FUNCTION_BLOCK MOD_StateLatch (* Keeps the last module state heard on the state channel. Technical: Local channel IDs of the PackML state and its refresh query; types and forwards the received PackML state *)
  (* Standard: 61499-2 *)
  (* Version 0.1, 2026-09-28, Project contributors, AAU Smart Production Lab *)
  PACKAGE modlib;
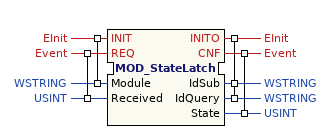
  EVENT_INPUT
    INIT : EInit WITH Module; (* Initialise, once at start-up (the INIT chain); takes the values given with it *)
    REQ WITH Received; (* The value arrived on the local channel *)
  END_EVENT
  EVENT_OUTPUT
    INITO : EInit WITH IdSub, IdQuery; (* Initialised: the next block of the INIT chain goes on *)
    CNF WITH State; (* Confirmation of REQ *)
  END_EVENT
  VAR_INPUT
    Module : WSTRING; (* The module's name; its local channels are named after it (loc[<Module>/...]) *)
    Received : USINT; (* The value as it arrived *)
  END_VAR
  VAR_OUTPUT
    IdSub : WSTRING; (* Local channel the value arrives on *)
    IdQuery : WSTRING; (* Local channel that asks for the current value (a block that starts later) *)
    State : USINT; (* PackML state: 1 Clearing, 2 Stopped, 3 Starting, 4 Idle, 6 Execute, 7 Stopping, 8 Aborting, 9 Aborted, 15 Resetting *)
  END_VAR
  EC_STATES
    INIT : INIT -> INITO;
    REQ : REQ -> CNF;
  END_STATES
  ALGORITHM INIT IN ST:
IdSub := CONCAT(CONCAT("loc[", Module), "/state]");
IdQuery := CONCAT(CONCAT("loc[", Module), "/state/query]");
  END_ALGORITHM
  ALGORITHM REQ IN ST:
State := Received;
  END_ALGORITHM
END_FUNCTION_BLOCK
